(* IEC 61131-3 sources: plc-st-coding-agent/progress/evidence/f14_v3_parallel_20261112/jobs/codex_minimax-m27 (part 3) *)

(* ---- self-hard-01.raw_candidate_02.st ---- *)
FUNCTION_BLOCK FB
VAR_INPUT
    flowLow   : BOOL;
    ackBtn    : BOOL;
    sensorOK  : BOOL;
END_VAR
VAR_OUTPUT
    alarmActive : BOOL;
    alarmAcked  : BOOL;
    highHigh    : BOOL;
END_VAR
VAR
    prev_flowLow : BOOL := FALSE;
    prev_ackBtn  : BOOL := FALSE;
END_VAR

VAR_TEMP
    risingAck : BOOL;
END_VAR

risingAck := ackBtn AND NOT prev_ackBtn;

IF flowLow THEN
    // Condition is active
    IF NOT alarmActive THEN
        // New alarm activation
        alarmActive := TRUE;
        alarmAcked  := FALSE;
    ELSIF risingAck THEN
        // Rising ack while condition still exists - just mark acknowledged
        alarmAcked := TRUE;
    END_IF;
ELSE
    // Condition has disappeared
    IF prev_flowLow AND alarmAcked THEN
        // Condition just cleared, was already acknowledged - clear immediately
        alarmActive := FALSE;
        alarmAcked  := FALSE;
    ELSIF prev_flowLow AND NOT alarmAcked THEN
        // Condition just cleared, unacknowledged - enter pending clear state
        alarmAcked := TRUE;
    ELSIF risingAck AND alarmAcked THEN
        // Condition still gone from before, pending clear - clear on new ack
        alarmActive := FALSE;
        alarmAcked  := FALSE;
    END_IF;
END_IF;

// High priority alarm: sensor failure (independent)
highHigh := NOT sensorOK;

// Update state for next cycle
prev_flowLow := flowLow;
prev_ackBtn  := ackBtn;

END_FUNCTION_BLOCK

(* ---- self-hard-02.candidate_01.st ---- *)
FUNCTION_BLOCK FB
VAR_INPUT
    startBtn    : BOOL;
    abortBtn    : BOOL;
    setpoint    : REAL;
    pv          : REAL;
    maxDuration : INT;
END_VAR
VAR_OUTPUT
    elapsed : INT := 0;
    phase   : INT := 0;
    timeout : BOOL := FALSE;
END_VAR
VAR
    prev_startBtn : BOOL := FALSE;
    prev_phase    : INT  := 0;
    prev_elapsed  : INT  := 0;
    prev_timeout  : BOOL := FALSE;
END_VAR

// Priority 1: Abort (highest)
IF abortBtn THEN
    phase   := 9;
    elapsed := prev_elapsed;
    timeout := prev_timeout;

// Priority 2: New start rising edge (no abort)
ELSIF startBtn AND NOT prev_startBtn THEN
    phase   := 1;
    elapsed := 0;
    timeout := FALSE;

// Priority 3: Running states (prev phase 1 or 2)
ELSIF prev_phase = 1 OR prev_phase = 2 THEN
    elapsed := prev_elapsed + 1;

    IF elapsed >= maxDuration THEN
        timeout := TRUE;
        phase   := 3;
    ELSIF prev_phase = 1 AND pv >= setpoint THEN
        phase := 2;
    ELSE
        phase := prev_phase;
    END_IF;

// Priority 4: Frozen states (phase 0, 3, 9)
ELSE
    phase   := prev_phase;
    elapsed := prev_elapsed;
    timeout := prev_timeout;
END_IF;

prev_startBtn := startBtn;
prev_phase    := phase;
prev_elapsed  := elapsed;
prev_timeout  := timeout;
END_FUNCTION_BLOCK

(* ---- self-hard-02.raw_candidate_01.st ---- *)
FUNCTION_BLOCK FB
VAR_INPUT
    startBtn    : BOOL;
    abortBtn    : BOOL;
    setpoint    : REAL;
    pv          : REAL;
    maxDuration : INT;
END_VAR
VAR_OUTPUT
    elapsed : INT := 0;
    phase   : INT := 0;
    timeout : BOOL := FALSE;
END_VAR
VAR
    prev_startBtn : BOOL := FALSE;
    prev_phase    : INT  := 0;
    prev_elapsed  : INT  := 0;
    prev_timeout  : BOOL := FALSE;
END_VAR

// Priority 1: Abort (highest)
IF abortBtn THEN
    phase   := 9;
    elapsed := prev_elapsed;
    timeout := prev_timeout;

// Priority 2: New start rising edge (no abort)
ELSIF startBtn AND NOT prev_startBtn THEN
    phase   := 1;
    elapsed := 0;
    timeout := FALSE;

// Priority 3: Running states (prev phase 1 or 2)
ELSIF prev_phase = 1 OR prev_phase = 2 THEN
    elapsed := prev_elapsed + 1;

    IF elapsed >= maxDuration THEN
        timeout := TRUE;
        phase   := 3;
    ELSIF prev_phase = 1 AND pv >= setpoint THEN
        phase := 2;
    ELSE
        phase := prev_phase;
    END_IF;

// Priority 4: Frozen states (phase 0, 3, 9)
ELSE
    phase   := prev_phase;
    elapsed := prev_elapsed;
    timeout := prev_timeout;
END_IF;

prev_startBtn := startBtn;
prev_phase    := phase;
prev_elapsed  := elapsed;
prev_timeout  := timeout;
END_FUNCTION_BLOCK

(* ---- self-hard-03.candidate_01.st ---- *)
FUNCTION_BLOCK FB
VAR_INPUT
    pushEn: BOOL;
    pushItem: INT;
    popEn: BOOL;
END_VAR

VAR_IN_OUT
    fifo: ARRAY[1..8] OF INT;
END_VAR

VAR_OUTPUT
    count: INT := 0;
    full: BOOL := FALSE;
    empty: BOOL := TRUE;
    head: INT := 0;
END_VAR

VAR
    prevPushEn: BOOL := FALSE;
    prevPopEn: BOOL := FALSE;
END_VAR

VAR
    risingPush: BOOL;
    risingPop: BOOL;
    i: INT;
END_VAR

// Detect rising edges
risingPush := pushEn AND NOT prevPushEn;
risingPop := popEn AND NOT prevPopEn;

// Process in order: pop first, then push
// POP: only if queue not empty
IF risingPop AND count > 0 THEN
    // Shift left if more than one element
    IF count > 1 THEN
        FOR i := 1 TO count - 1 DO
            fifo[i] := fifo[i + 1];
        END_FOR;
    END_IF;
    // Decrement count
    count := count - 1;
END_IF;

// PUSH: only if queue not full
IF risingPush AND count < 8 THEN
    count := count + 1;
    fifo[count] := pushItem;
END_IF;

// Update outputs
full := (count = 8);
empty := (count = 0);
IF count > 0 THEN
    head := fifo[1];
ELSE
    head := 0;
END_IF;

// Save current state for next cycle
prevPushEn := pushEn;
prevPopEn := popEn;

END_FUNCTION_BLOCK

(* ---- self-hard-03.raw_candidate_01.st ---- *)
FUNCTION_BLOCK FB
VAR_INPUT
    pushEn: BOOL;
    pushItem: INT;
    popEn: BOOL;
END_VAR

VAR_IN_OUT
    fifo: ARRAY[1..8] OF INT;
END_VAR

VAR_OUTPUT
    count: INT := 0;
    full: BOOL := FALSE;
    empty: BOOL := TRUE;
    head: INT := 0;
END_VAR

VAR
    prevPushEn: BOOL := FALSE;
    prevPopEn: BOOL := FALSE;
END_VAR

VAR
    risingPush: BOOL;
    risingPop: BOOL;
    i: INT;
END_VAR

// Detect rising edges
risingPush := pushEn AND NOT prevPushEn;
risingPop := popEn AND NOT prevPopEn;

// Process in order: pop first, then push
// POP: only if queue not empty
IF risingPop AND count > 0 THEN
    // Shift left if more than one element
    IF count > 1 THEN
        FOR i := 1 TO count - 1 DO
            fifo[i] := fifo[i + 1];
        END_FOR;
    END_IF;
    // Decrement count
    count := count - 1;
END_IF;

// PUSH: only if queue not full
IF risingPush AND count < 8 THEN
    count := count + 1;
    fifo[count] := pushItem;
END_IF;

// Update outputs
full := (count = 8);
empty := (count = 0);
IF count > 0 THEN
    head := fifo[1];
ELSE
    head := 0;
END_IF;

// Save current state for next cycle
prevPushEn := pushEn;
prevPopEn := popEn;

END_FUNCTION_BLOCK

(* ---- self-hard-04.candidate_01.st ---- *)
FUNCTION_BLOCK FB
VAR
    prevDemand: INT := 0;
    prevLeadPump: INT := 0;
    prevRunningCount: INT := 0;
    prevLagPump: INT := 0;
    leadPump: INT := 0;
    lagPump: INT := 0;
    runningCount: INT := 0;
    minHours: LINT;
    minPumpIdx: INT;
    secondMinHours: LINT;
    secondMinIdx: INT;
    hoursDiff: LINT;
    needInitialLead: BOOL;
    needSwitchLead: BOOL;
    needRefreshLag: BOOL;
    i: INT;
    h: LINT;
END_VAR

// Clip demand to 0..5
IF demand < 0 THEN
    runningCount := 0;
ELSIF demand > 5 THEN
    runningCount := 5;
ELSE
    runningCount := demand;
END_IF;

// Detect state transitions
needInitialLead := (prevDemand = 0) AND (runningCount > 0);
needRefreshLag := (runningCount > prevRunningCount) OR (leadPump <> prevLeadPump);

// Find pump with minimum (runHours, pumpIdx)
minHours := runHours[1];
minPumpIdx := 1;
FOR i := 2 TO 5 DO
    h := runHours[i];
    IF (h < minHours) OR ((h = minHours) AND (i < minPumpIdx)) THEN
        minHours := h;
        minPumpIdx := i;
    END_IF;
END_FOR;

// Lead pump hysteresis check
IF leadPump >= 1 AND leadPump <= 5 THEN
    hoursDiff := runHours[leadPump] - minHours;
ELSE
    hoursDiff := 0;
END_IF;
needSwitchLead := (prevLeadPump <> 0) AND rotated AND (hoursDiff > 50);

// Demand = 0: clear both pumps immediately
IF runningCount = 0 THEN
    leadPump := 0;
    lagPump := 0;
    needRefreshLag := FALSE;
    needSwitchLead := FALSE;
END_IF;

// Handle lead pump change
IF needSwitchLead THEN
    leadPump := minPumpIdx;
    needRefreshLag := TRUE;
ELSIF needInitialLead THEN
    leadPump := minPumpIdx;
END_IF;

// Lag pump selection
IF needRefreshLag AND runningCount > 0 THEN
    secondMinHours := 16#7FFFFFFFFFFFFFFF;
    secondMinIdx := 0;
    FOR i := 1 TO 5 DO
        IF i <> leadPump THEN
            h := runHours[i];
            IF (h < secondMinHours) OR ((h = secondMinHours) AND (i < secondMinIdx)) THEN
                secondMinHours := h;
                secondMinIdx := i;
            END_IF;
        END_IF;
    END_FOR;
    lagPump := secondMinIdx;
ELSIF runningCount = 1 THEN
    lagPump := 0;
END_IF;

// Preserve lead pump if no change occurred
IF NOT needSwitchLead AND NOT needInitialLead AND runningCount > 0 THEN
    leadPump := prevLeadPump;
END_IF;

// Update previous-cycle state
prevDemand := runningCount;
prevLeadPump := leadPump;
prevRunningCount := runningCount;
prevLagPump := lagPump;

END_FUNCTION_BLOCK

(* ---- self-hard-04.candidate_02.st ---- *)
FUNCTION_BLOCK FB
VAR_INPUT
    demand: INT;
    runHours: ARRAY[1..5] OF LINT;
    rotated: BOOL;
END_VAR
VAR_OUTPUT
    leadPump: INT;
    lagPump: INT;
    runningCount: INT;
END_VAR
VAR
    prevDemand: INT := 0;
    prevLeadPump: INT := 0;
    prevRunningCount: INT := 0;
    prevLagPump: INT := 0;
    minHours: LINT;
    minPumpIdx: INT;
    secondMinHours: LINT;
    secondMinIdx: INT;
    hoursDiff: LINT;
    needInitialLead: BOOL;
    needSwitchLead: BOOL;
    needRefreshLag: BOOL;
    i: INT;
    h: LINT;
    clippedDemand: INT;
END_VAR

clippedDemand := demand;
IF clippedDemand < 0 THEN
    clippedDemand := 0;
ELSIF clippedDemand > 5 THEN
    clippedDemand := 5;
END_IF;

runningCount := clippedDemand;

needInitialLead := (prevDemand = 0) AND (runningCount > 0);
needRefreshLag := (runningCount > prevRunningCount) OR (leadPump <> prevLeadPump);

minHours := runHours[1];
minPumpIdx := 1;
FOR i := 2 TO 5 DO
    h := runHours[i];
    IF (h < minHours) OR ((h = minHours) AND (i < minPumpIdx)) THEN
        minHours := h;
        minPumpIdx := i;
    END_IF;
END_FOR;

IF leadPump >= 1 AND leadPump <= 5 THEN
    hoursDiff := runHours[leadPump] - minHours;
ELSE
    hoursDiff := 0;
END_IF;

needSwitchLead := (prevLeadPump <> 0) AND rotated AND (hoursDiff > 50);

IF runningCount = 0 THEN
    leadPump := 0;
    lagPump := 0;
ELSIF needSwitchLead THEN
    leadPump := minPumpIdx;
ELSIF needInitialLead THEN
    leadPump := minPumpIdx;
ELSE
    leadPump := prevLeadPump;
END_IF;

IF runningCount >= 2 THEN
    IF needRefreshLag THEN
        secondMinHours := 16#7FFFFFFFFFFFFFFF;
        secondMinIdx := 0;
        FOR i := 1 TO 5 DO
            IF i <> leadPump THEN
                h := runHours[i];
                IF (h < secondMinHours) OR ((h = secondMinHours) AND (i < secondMinIdx)) THEN
                    secondMinHours := h;
                    secondMinIdx := i;
                END_IF;
            END_IF;
        END_FOR;
        lagPump := secondMinIdx;
    ELSE
        lagPump := prevLagPump;
    END_IF;
ELSE
    lagPump := 0;
END_IF;

prevDemand := clippedDemand;
prevLeadPump := leadPump;
prevRunningCount := runningCount;
prevLagPump := lagPump;

END_FUNCTION_BLOCK

(* ---- self-hard-04.raw_candidate_01.st ---- *)
FUNCTION_BLOCK FB
VAR
    prevDemand: INT := 0;
    prevLeadPump: INT := 0;
    prevRunningCount: INT := 0;
    prevLagPump: INT := 0;
    leadPump: INT := 0;
    lagPump: INT := 0;
    runningCount: INT := 0;
    minHours: LINT;
    minPumpIdx: INT;
    secondMinHours: LINT;
    secondMinIdx: INT;
    hoursDiff: LINT;
    needInitialLead: BOOL;
    needSwitchLead: BOOL;
    needRefreshLag: BOOL;
    i: INT;
    h: LINT;
END_VAR

// Clip demand to 0..5
IF demand < 0 THEN
    runningCount := 0;
ELSIF demand > 5 THEN
    runningCount := 5;
ELSE
    runningCount := demand;
END_IF;

// Detect state transitions
needInitialLead := (prevDemand = 0) AND (runningCount > 0);
needRefreshLag := (runningCount > prevRunningCount) OR (leadPump <> prevLeadPump);

// Find pump with minimum (runHours, pumpIdx)
minHours := runHours[1];
minPumpIdx := 1;
FOR i := 2 TO 5 DO
    h := runHours[i];
    IF (h < minHours) OR ((h = minHours) AND (i < minPumpIdx)) THEN
        minHours := h;
        minPumpIdx := i;
    END_IF;
END_FOR;

// Lead pump hysteresis check
IF leadPump >= 1 AND leadPump <= 5 THEN
    hoursDiff := runHours[leadPump] - minHours;
ELSE
    hoursDiff := 0;
END_IF;
needSwitchLead := (prevLeadPump <> 0) AND rotated AND (hoursDiff > 50);

// Demand = 0: clear both pumps immediately
IF runningCount = 0 THEN
    leadPump := 0;
    lagPump := 0;
    needRefreshLag := FALSE;
    needSwitchLead := FALSE;
END_IF;

// Handle lead pump change
IF needSwitchLead THEN
    leadPump := minPumpIdx;
    needRefreshLag := TRUE;
ELSIF needInitialLead THEN
    leadPump := minPumpIdx;
END_IF;

// Lag pump selection
IF needRefreshLag AND runningCount > 0 THEN
    secondMinHours := 16#7FFFFFFFFFFFFFFF;
    secondMinIdx := 0;
    FOR i := 1 TO 5 DO
        IF i <> leadPump THEN
            h := runHours[i];
            IF (h < secondMinHours) OR ((h = secondMinHours) AND (i < secondMinIdx)) THEN
                secondMinHours := h;
                secondMinIdx := i;
            END_IF;
        END_IF;
    END_FOR;
    lagPump := secondMinIdx;
ELSIF runningCount = 1 THEN
    lagPump := 0;
END_IF;

// Preserve lead pump if no change occurred
IF NOT needSwitchLead AND NOT needInitialLead AND runningCount > 0 THEN
    leadPump := prevLeadPump;
END_IF;

// Update previous-cycle state
prevDemand := runningCount;
prevLeadPump := leadPump;
prevRunningCount := runningCount;
prevLagPump := lagPump;

END_FUNCTION_BLOCK

(* ---- self-hard-04.raw_candidate_02.st ---- *)
FUNCTION_BLOCK FB
VAR_INPUT
    demand: INT;
    runHours: ARRAY[1..5] OF LINT;
    rotated: BOOL;
END_VAR
VAR_OUTPUT
    leadPump: INT;
    lagPump: INT;
    runningCount: INT;
END_VAR
VAR
    prevDemand: INT := 0;
    prevLeadPump: INT := 0;
    prevRunningCount: INT := 0;
    prevLagPump: INT := 0;
    minHours: LINT;
    minPumpIdx: INT;
    secondMinHours: LINT;
    secondMinIdx: INT;
    hoursDiff: LINT;
    needInitialLead: BOOL;
    needSwitchLead: BOOL;
    needRefreshLag: BOOL;
    i: INT;
    h: LINT;
    clippedDemand: INT;
END_VAR

clippedDemand := demand;
IF clippedDemand < 0 THEN
    clippedDemand := 0;
ELSIF clippedDemand > 5 THEN
    clippedDemand := 5;
END_IF;

runningCount := clippedDemand;

needInitialLead := (prevDemand = 0) AND (runningCount > 0);
needRefreshLag := (runningCount > prevRunningCount) OR (leadPump <> prevLeadPump);

minHours := runHours[1];
minPumpIdx := 1;
FOR i := 2 TO 5 DO
    h := runHours[i];
    IF (h < minHours) OR ((h = minHours) AND (i < minPumpIdx)) THEN
        minHours := h;
        minPumpIdx := i;
    END_IF;
END_FOR;

IF leadPump >= 1 AND leadPump <= 5 THEN
    hoursDiff := runHours[leadPump] - minHours;
ELSE
    hoursDiff := 0;
END_IF;

needSwitchLead := (prevLeadPump <> 0) AND rotated AND (hoursDiff > 50);

IF runningCount = 0 THEN
    leadPump := 0;
    lagPump := 0;
ELSIF needSwitchLead THEN
    leadPump := minPumpIdx;
ELSIF needInitialLead THEN
    leadPump := minPumpIdx;
ELSE
    leadPump := prevLeadPump;
END_IF;

IF runningCount >= 2 THEN
    IF needRefreshLag THEN
        secondMinHours := 16#7FFFFFFFFFFFFFFF;
        secondMinIdx := 0;
        FOR i := 1 TO 5 DO
            IF i <> leadPump THEN
                h := runHours[i];
                IF (h < secondMinHours) OR ((h = secondMinHours) AND (i < secondMinIdx)) THEN
                    secondMinHours := h;
                    secondMinIdx := i;
                END_IF;
            END_IF;
        END_FOR;
        lagPump := secondMinIdx;
    ELSE
        lagPump := prevLagPump;
    END_IF;
ELSE
    lagPump := 0;
END_IF;

prevDemand := clippedDemand;
prevLeadPump := leadPump;
prevRunningCount := runningCount;
prevLagPump := lagPump;

END_FUNCTION_BLOCK

(* ---- self-hard-05.candidate_01.st ---- *)
FUNCTION_BLOCK FB
VAR_INPUT
    runRequest  : BOOL;
    flameOK     : BOOL;
    o2Valid     : BOOL;
    o2PV        : REAL;
    baseAir     : REAL;
    resetBtn    : BOOL;
END_VAR

VAR_OUTPUT
    fuelPermit  : BOOL;
    trimEnable  : BOOL;
    airTrim     : REAL;
    airCommand  : REAL;
    tripLatched : BOOL;
    o2Fault     : BOOL;
END_VAR

VAR
    prevResetBtn : BOOL := FALSE;
    tripInternal : BOOL := FALSE;
END_VAR

// 氧量故障判定
o2Fault := NOT o2Valid OR o2PV < 0.0 OR o2PV > 21.0;

// 熄火跳闸逻辑：运行中失去火焰当拍置位；安全停机态下复位上升沿清除
IF runRequest AND NOT flameOK THEN
    tripInternal := TRUE;
ELSIF NOT runRequest AND NOT flameOK AND resetBtn AND NOT prevResetBtn THEN
    tripInternal := FALSE;
END_IF;

// 燃料许可：运行请求、火焰正常、未跳闸三者同时成立
fuelPermit := runRequest AND flameOK AND NOT tripInternal;

// 氧量修正：投入需燃料许可且分析仪无故障
trimEnable := fuelPermit AND NOT o2Fault;
airTrim := 2.0 * (2.0 - o2PV);
airTrim := LIMIT(-10.0, airTrim, 10.0);
airTrim := SEL(trimEnable, 0.0, airTrim);

// 风门命令：基础开度叠加修正，偏置切除时自动归零
airCommand := baseAir + airTrim;
airCommand := LIMIT(0.0, airCommand, 100.0);
airCommand := SEL(fuelPermit, 0.0, airCommand);

// 输出跳闸状态
tripLatched := tripInternal;

// 边沿检测：保存复位按钮上一拍状态
prevResetBtn := resetBtn;

END_FUNCTION_BLOCK

(* ---- self-hard-05.candidate_02.st ---- *)
FUNCTION_BLOCK FB
VAR_INPUT
    runRequest  : BOOL;
    flameOK     : BOOL;
    o2Valid     : BOOL;
    o2PV        : REAL;
    baseAir     : REAL;
    resetBtn    : BOOL;
END_VAR

VAR_OUTPUT
    fuelPermit  : BOOL;
    trimEnable  : BOOL;
    airTrim     : REAL;
    airCommand  : REAL;
    tripLatched : BOOL;
    o2Fault     : BOOL;
END_VAR

VAR
    prevResetBtn : BOOL := FALSE;
    tripInternal : BOOL := FALSE;
END_VAR

// 氧量故障判定
o2Fault := NOT o2Valid OR o2PV < 0.0 OR o2PV > 21.0;

// 熄火跳闸逻辑：运行中失去火焰当拍置位；安全停机态下复位上升沿清除
IF runRequest AND NOT flameOK THEN
    tripInternal := TRUE;
ELSIF NOT runRequest AND NOT flameOK AND resetBtn AND NOT prevResetBtn THEN
    tripInternal := FALSE;
END_IF;

// 燃料许可：运行请求、火焰正常、未跳闸三者同时成立
fuelPermit := runRequest AND flameOK AND NOT tripInternal;

// 氧量修正：投入需燃料许可且分析仪无故障
IF fuelPermit AND NOT o2Fault THEN
    trimEnable := TRUE;
    airTrim := LIMIT(-10.0, 2.0 * (2.0 - o2PV), 10.0);
ELSE
    trimEnable := FALSE;
    airTrim := 0.0;
END_IF;

// 风门命令：基础开度叠加修正，偏置切除时自动归零
IF fuelPermit THEN
    airCommand := LIMIT(0.0, baseAir + airTrim, 100.0);
ELSE
    airCommand := 0.0;
END_IF;

// 输出跳闸状态
tripLatched := tripInternal;

// 边沿检测：保存复位按钮上一拍状态
prevResetBtn := resetBtn;

END_FUNCTION_BLOCK

(* ---- self-hard-05.raw_candidate_01.st ---- *)
FUNCTION_BLOCK FB
VAR_INPUT
    runRequest  : BOOL;
    flameOK     : BOOL;
    o2Valid     : BOOL;
    o2PV        : REAL;
    baseAir     : REAL;
    resetBtn    : BOOL;
END_VAR

VAR_OUTPUT
    fuelPermit  : BOOL;
    trimEnable  : BOOL;
    airTrim     : REAL;
    airCommand  : REAL;
    tripLatched : BOOL;
    o2Fault     : BOOL;
END_VAR

VAR
    prevResetBtn : BOOL := FALSE;
    tripInternal : BOOL := FALSE;
END_VAR

// 氧量故障判定
o2Fault := NOT o2Valid OR o2PV < 0.0 OR o2PV > 21.0;

// 熄火跳闸逻辑：运行中失去火焰当拍置位；安全停机态下复位上升沿清除
IF runRequest AND NOT flameOK THEN
    tripInternal := TRUE;
ELSIF NOT runRequest AND NOT flameOK AND resetBtn AND NOT prevResetBtn THEN
    tripInternal := FALSE;
END_IF;

// 燃料许可：运行请求、火焰正常、未跳闸三者同时成立
fuelPermit := runRequest AND flameOK AND NOT tripInternal;

// 氧量修正：投入需燃料许可且分析仪无故障
trimEnable := fuelPermit AND NOT o2Fault;
airTrim := 2.0 * (2.0 - o2PV);
airTrim := LIMIT(-10.0, airTrim, 10.0);
airTrim := SEL(trimEnable, 0.0, airTrim);

// 风门命令：基础开度叠加修正，偏置切除时自动归零
airCommand := baseAir + airTrim;
airCommand := LIMIT(0.0, airCommand, 100.0);
airCommand := SEL(fuelPermit, 0.0, airCommand);

// 输出跳闸状态
tripLatched := tripInternal;

// 边沿检测：保存复位按钮上一拍状态
prevResetBtn := resetBtn;

END_FUNCTION_BLOCK

(* ---- self-hard-05.raw_candidate_02.st ---- *)
FUNCTION_BLOCK FB
VAR_INPUT
    runRequest  : BOOL;
    flameOK     : BOOL;
    o2Valid     : BOOL;
    o2PV        : REAL;
    baseAir     : REAL;
    resetBtn    : BOOL;
END_VAR

VAR_OUTPUT
    fuelPermit  : BOOL;
    trimEnable  : BOOL;
    airTrim     : REAL;
    airCommand  : REAL;
    tripLatched : BOOL;
    o2Fault     : BOOL;
END_VAR

VAR
    prevResetBtn : BOOL := FALSE;
    tripInternal : BOOL := FALSE;
END_VAR

// 氧量故障判定
o2Fault := NOT o2Valid OR o2PV < 0.0 OR o2PV > 21.0;

// 熄火跳闸逻辑：运行中失去火焰当拍置位；安全停机态下复位上升沿清除
IF runRequest AND NOT flameOK THEN
    tripInternal := TRUE;
ELSIF NOT runRequest AND NOT flameOK AND resetBtn AND NOT prevResetBtn THEN
    tripInternal := FALSE;
END_IF;

// 燃料许可：运行请求、火焰正常、未跳闸三者同时成立
fuelPermit := runRequest AND flameOK AND NOT tripInternal;

// 氧量修正：投入需燃料许可且分析仪无故障
IF fuelPermit AND NOT o2Fault THEN
    trimEnable := TRUE;
    airTrim := LIMIT(-10.0, 2.0 * (2.0 - o2PV), 10.0);
ELSE
    trimEnable := FALSE;
    airTrim := 0.0;
END_IF;

// 风门命令：基础开度叠加修正，偏置切除时自动归零
IF fuelPermit THEN
    airCommand := LIMIT(0.0, baseAir + airTrim, 100.0);
ELSE
    airCommand := 0.0;
END_IF;

// 输出跳闸状态
tripLatched := tripInternal;

// 边沿检测：保存复位按钮上一拍状态
prevResetBtn := resetBtn;

END_FUNCTION_BLOCK

(* ---- self-hard-06.candidate_01.st ---- *)
FUNCTION_BLOCK FB
VAR_INPUT
    runRequest      : BOOL;
    pressure        : REAL;
    pressureValid   : BOOL;
    fuelFlow        : REAL;
    steamFlow       : REAL;
    outletCmd       : INT;
    outletFeedback  : INT;
    resetBtn        : BOOL;
END_VAR
VAR_OUTPUT
    tripLatched     : BOOL;
    fuelPermit      : BOOL;
    currentCauseMask: WORD;
    latchedCauseMask: WORD;
    diagnosticActive: BOOL;
END_VAR
VAR
    prevResetBtn    : BOOL := FALSE;
    stickyCounter   : INT  := 0;
END_VAR

// Reset edge detection
IF resetBtn AND NOT prevResetBtn THEN
    // Rising edge of reset button
    IF NOT runRequest AND pressureValid AND pressure <= 4200.0 THEN
        tripLatched     := FALSE;
        latchedCauseMask := 0;
    ELSE
        tripLatched := TRUE;
    END_IF;
ELSE
    // No reset edge
    IF tripLatched THEN
        tripLatched := TRUE;
    ELSIF runRequest AND (NOT pressureValid OR pressure >= 4500.0) THEN
        tripLatched := TRUE;
    END_IF;
END_IF;

// Valve sticking counter: reset on any interruption, increment only in valid overpressure
IF NOT runRequest OR NOT pressureValid OR pressure < 4500.0 OR outletCmd < 50 OR outletFeedback > 10 THEN
    stickyCounter := 0;
ELSIF outletCmd >= 50 AND outletFeedback <= 10 THEN
    stickyCounter := stickyCounter + 1;
END_IF;

// Determine current cause mask
currentCauseMask := 0;
IF runRequest THEN
    IF NOT pressureValid THEN
        currentCauseMask := 1;  // bit0 = 1
    ELSIF stickyCounter >= 3 THEN
        currentCauseMask := 2;  // bit1 = 2
    END_IF;

    IF pressureValid AND pressure >= 4500.0 THEN
        IF fuelFlow >= 4.0 AND steamFlow <= 10.0 THEN
            currentCauseMask := currentCauseMask OR 4;  // bit2 = 4
        END_IF;

        IF currentCauseMask = 0 THEN
            currentCauseMask := 8;  // bit3 = 8
        END_IF;
    END_IF;
END_IF;

// Accumulate latched mask during trip
IF tripLatched THEN
    latchedCauseMask := latchedCauseMask OR currentCauseMask;
END_IF;

// Outputs
fuelPermit      := runRequest AND NOT tripLatched;
diagnosticActive := (currentCauseMask <> 0);

// Update previous states
prevResetBtn := resetBtn;
END_FUNCTION_BLOCK

(* ---- self-hard-06.candidate_02.st ---- *)
FUNCTION_BLOCK FB
VAR_INPUT
    runRequest       : BOOL;
    pressure         : REAL;
    pressureValid    : BOOL;
    fuelFlow         : REAL;
    steamFlow        : REAL;
    outletCmd        : INT;
    outletFeedback   : INT;
    resetBtn         : BOOL;
END_VAR
VAR_OUTPUT
    tripLatched      : BOOL;
    fuelPermit       : BOOL;
    currentCauseMask : WORD;
    latchedCauseMask : WORD;
    diagnosticActive : BOOL;
END_VAR
VAR
    prevResetBtn     : BOOL := FALSE;
    stickyCounter    : INT  := 0;
END_VAR

// Rising edge detection for reset
VAR_TEMP
    resetRising : BOOL;
END_VAR
resetRising := resetBtn AND NOT prevResetBtn;

// S17 logic: latch holds from first trip until valid reset edge
IF resetRising AND NOT runRequest AND pressureValid AND pressure <= 4200.0 THEN
    tripLatched := FALSE;
    latchedCauseMask := 0;
ELSIF resetRising THEN
    tripLatched := TRUE;
    IF tripLatched THEN
        latchedCauseMask := latchedCauseMask OR currentCauseMask;
    END_IF;
ELSIF prevResetBtn OR tripLatched THEN
    tripLatched := TRUE;
    IF prevResetBtn OR tripLatched THEN
        latchedCauseMask := latchedCauseMask OR currentCauseMask;
    END_IF;
ELSIF runRequest AND (NOT pressureValid OR pressure >= 4500.0) THEN
    tripLatched := TRUE;
    latchedCauseMask := currentCauseMask;
ELSE
    tripLatched := FALSE;
END_IF;

// Valve sticking counter
IF NOT runRequest OR NOT pressureValid OR pressure < 4500.0 OR outletCmd < 50 OR outletFeedback > 10 THEN
    stickyCounter := 0;
ELSIF outletCmd >= 50 AND outletFeedback <= 10 THEN
    stickyCounter := stickyCounter + 1;
END_IF;

// Current cause mask
currentCauseMask := 0;
IF runRequest THEN
    IF NOT pressureValid THEN
        currentCauseMask := 1;
    ELSIF stickyCounter >= 3 THEN
        currentCauseMask := 2;
    END_IF;

    IF pressureValid AND pressure >= 4500.0 THEN
        IF fuelFlow >= 4.0 AND steamFlow <= 10.0 THEN
            currentCauseMask := currentCauseMask OR 4;
        END_IF;

        IF currentCauseMask = 0 THEN
            currentCauseMask := 8;
        END_IF;
    END_IF;
END_IF;

// Outputs
fuelPermit       := runRequest AND NOT tripLatched;
diagnosticActive := (currentCauseMask <> 0);

prevResetBtn := resetBtn;
END_FUNCTION_BLOCK

(* ---- self-hard-06.raw_candidate_01.st ---- *)
FUNCTION_BLOCK FB
VAR_INPUT
    runRequest      : BOOL;
    pressure        : REAL;
    pressureValid   : BOOL;
    fuelFlow        : REAL;
    steamFlow       : REAL;
    outletCmd       : INT;
    outletFeedback  : INT;
    resetBtn        : BOOL;
END_VAR
VAR_OUTPUT
    tripLatched     : BOOL;
    fuelPermit      : BOOL;
    currentCauseMask: WORD;
    latchedCauseMask: WORD;
    diagnosticActive: BOOL;
END_VAR
VAR
    prevResetBtn    : BOOL := FALSE;
    stickyCounter   : INT  := 0;
END_VAR

// Reset edge detection
IF resetBtn AND NOT prevResetBtn THEN
    // Rising edge of reset button
    IF NOT runRequest AND pressureValid AND pressure <= 4200.0 THEN
        tripLatched     := FALSE;
        latchedCauseMask := 0;
    ELSE
        tripLatched := TRUE;
    END_IF;
ELSE
    // No reset edge
    IF tripLatched THEN
        tripLatched := TRUE;
    ELSIF runRequest AND (NOT pressureValid OR pressure >= 4500.0) THEN
        tripLatched := TRUE;
    END_IF;
END_IF;

// Valve sticking counter: reset on any interruption, increment only in valid overpressure
IF NOT runRequest OR NOT pressureValid OR pressure < 4500.0 OR outletCmd < 50 OR outletFeedback > 10 THEN
    stickyCounter := 0;
ELSIF outletCmd >= 50 AND outletFeedback <= 10 THEN
    stickyCounter := stickyCounter + 1;
END_IF;

// Determine current cause mask
currentCauseMask := 0;
IF runRequest THEN
    IF NOT pressureValid THEN
        currentCauseMask := 1;  // bit0 = 1
    ELSIF stickyCounter >= 3 THEN
        currentCauseMask := 2;  // bit1 = 2
    END_IF;

    IF pressureValid AND pressure >= 4500.0 THEN
        IF fuelFlow >= 4.0 AND steamFlow <= 10.0 THEN
            currentCauseMask := currentCauseMask OR 4;  // bit2 = 4
        END_IF;

        IF currentCauseMask = 0 THEN
            currentCauseMask := 8;  // bit3 = 8
        END_IF;
    END_IF;
END_IF;

// Accumulate latched mask during trip
IF tripLatched THEN
    latchedCauseMask := latchedCauseMask OR currentCauseMask;
END_IF;

// Outputs
fuelPermit      := runRequest AND NOT tripLatched;
diagnosticActive := (currentCauseMask <> 0);

// Update previous states
prevResetBtn := resetBtn;
END_FUNCTION_BLOCK

(* ---- self-hard-06.raw_candidate_02.st ---- *)
FUNCTION_BLOCK FB
VAR_INPUT
    runRequest       : BOOL;
    pressure         : REAL;
    pressureValid    : BOOL;
    fuelFlow         : REAL;
    steamFlow        : REAL;
    outletCmd        : INT;
    outletFeedback   : INT;
    resetBtn         : BOOL;
END_VAR
VAR_OUTPUT
    tripLatched      : BOOL;
    fuelPermit       : BOOL;
    currentCauseMask : WORD;
    latchedCauseMask : WORD;
    diagnosticActive : BOOL;
END_VAR
VAR
    prevResetBtn     : BOOL := FALSE;
    stickyCounter    : INT  := 0;
END_VAR

// Rising edge detection for reset
VAR_TEMP
    resetRising : BOOL;
END_VAR
resetRising := resetBtn AND NOT prevResetBtn;

// S17 logic: latch holds from first trip until valid reset edge
IF resetRising AND NOT runRequest AND pressureValid AND pressure <= 4200.0 THEN
    tripLatched := FALSE;
    latchedCauseMask := 0;
ELSIF resetRising THEN
    tripLatched := TRUE;
    IF tripLatched THEN
        latchedCauseMask := latchedCauseMask OR currentCauseMask;
    END_IF;
ELSIF prevResetBtn OR tripLatched THEN
    tripLatched := TRUE;
    IF prevResetBtn OR tripLatched THEN
        latchedCauseMask := latchedCauseMask OR currentCauseMask;
    END_IF;
ELSIF runRequest AND (NOT pressureValid OR pressure >= 4500.0) THEN
    tripLatched := TRUE;
    latchedCauseMask := currentCauseMask;
ELSE
    tripLatched := FALSE;
END_IF;

// Valve sticking counter
IF NOT runRequest OR NOT pressureValid OR pressure < 4500.0 OR outletCmd < 50 OR outletFeedback > 10 THEN
    stickyCounter := 0;
ELSIF outletCmd >= 50 AND outletFeedback <= 10 THEN
    stickyCounter := stickyCounter + 1;
END_IF;

// Current cause mask
currentCauseMask := 0;
IF runRequest THEN
    IF NOT pressureValid THEN
        currentCauseMask := 1;
    ELSIF stickyCounter >= 3 THEN
        currentCauseMask := 2;
    END_IF;

    IF pressureValid AND pressure >= 4500.0 THEN
        IF fuelFlow >= 4.0 AND steamFlow <= 10.0 THEN
            currentCauseMask := currentCauseMask OR 4;
        END_IF;

        IF currentCauseMask = 0 THEN
            currentCauseMask := 8;
        END_IF;
    END_IF;
END_IF;

// Outputs
fuelPermit       := runRequest AND NOT tripLatched;
diagnosticActive := (currentCauseMask <> 0);

prevResetBtn := resetBtn;
END_FUNCTION_BLOCK

(* ---- self-hard-07.candidate_01.st ---- *)
FUNCTION_BLOCK FB
VAR_INPUT
    mode            : INT;
    resetBtn        : BOOL;
    scanSeconds     : REAL;
    tempSP          : REAL;
    tempPV          : REAL;
    flowPV          : REAL;
    manualFlowSP    : REAL;
    manualValve     : REAL;
END_VAR

VAR_OUTPUT
    flowSP          : REAL;
    valveCommand    : REAL;
    fault           : BOOL;
    normalMode      : BOOL;
END_VAR

VAR
    prevMode        : INT;
    prevResetBtn    : BOOL;
    prevFlowSP      : REAL;
    prevValveCmd    : REAL;
    prevTempSP      : REAL;
    accT            : REAL;
    accF            : REAL;
    firstScan       : BOOL;
END_VAR

fault := (mode < 0) OR (mode > 2) OR (scanSeconds <= 0.0) OR (scanSeconds > 10.0);

IF resetBtn AND NOT prevResetBtn THEN
    flowSP := manualFlowSP;
    valveCommand := manualValve;
    accT := 0.0;
    accF := 0.0;
    normalMode := FALSE;
    firstScan := FALSE;
    prevMode := mode;
    prevResetBtn := resetBtn;
    prevFlowSP := flowSP;
    prevValveCmd := valveCommand;
    prevTempSP := tempSP;
    RETURN;
END_IF;

IF mode <> prevMode THEN
    IF mode = 2 THEN
        flowSP := prevFlowSP;
        valveCommand := prevValveCmd;
    ELSE
        flowSP := manualFlowSP;
        valveCommand := prevValveCmd;
    END_IF;
    normalMode := FALSE;
    prevMode := mode;
    prevResetBtn := resetBtn;
    prevFlowSP := flowSP;
    prevValveCmd := valveCommand;
    prevTempSP := tempSP;
    RETURN;
END_IF;

IF firstScan THEN
    flowSP := manualFlowSP;
    valveCommand := manualValve;
    accT := 0.0;
    accF := 0.0;
    normalMode := FALSE;
    firstScan := FALSE;
    prevMode := mode;
    prevResetBtn := resetBtn;
    prevFlowSP := flowSP;
    prevValveCmd := valveCommand;
    prevTempSP := tempSP;
    RETURN;
END_IF;

normalMode := TRUE;

IF mode = 2 THEN
    VAR eF AT%Q* : REAL; END_VAR
    eF := flowSP - flowPV;
    accF := accF + 0.5 * eF * scanSeconds;
    valveCommand := 2.0 * eF + accF;
    valveCommand := LIMIT(0.0, valveCommand, 100.0);
    accF := valveCommand - 2.0 * eF;

    VAR eT AT%Q* : REAL; END_VAR
    eT := tempSP - tempPV;
    accT := accT + 0.2 * eT * scanSeconds;
    flowSP := 1.0 * eT + accT;
    flowSP := LIMIT(0.0, flowSP, 50.0);
    accT := flowSP - 1.0 * eT;
ELSIF mode = 1 THEN
    VAR eF AT%Q* : REAL; END_VAR
    eF := flowSP - flowPV;
    accF := accF + 0.5 * eF * scanSeconds;
    valveCommand := 2.0 * eF + accF;
    valveCommand := LIMIT(0.0, valveCommand, 100.0);
    accF := valveCommand - 2.0 * eF;
ELSE
    flowSP := manualFlowSP;
    valveCommand := manualValve;
END_IF;

prevMode := mode;
prevResetBtn := resetBtn;
prevFlowSP := flowSP;
prevValveCmd := valveCommand;
prevTempSP := tempSP;

END_FUNCTION_BLOCK

(* ---- self-hard-07.candidate_02.st ---- *)
FUNCTION_BLOCK FB
VAR_INPUT
    mode            : INT;
    resetBtn        : BOOL;
    scanSeconds     : REAL;
    tempSP          : REAL;
    tempPV          : REAL;
    flowPV          : REAL;
    manualFlowSP    : REAL;
    manualValve     : REAL;
END_VAR

VAR_OUTPUT
    flowSP          : REAL;
    valveCommand    : REAL;
    fault           : BOOL;
    normalMode      : BOOL;
END_VAR

VAR
    prevMode        : INT;
    prevResetBtn    : BOOL;
    prevFlowSP      : REAL;
    prevValveCmd    : REAL;
    accT            : REAL;
    accF            : REAL;
    firstScan       : BOOL;
    modeChanged     : BOOL;
END_VAR

    modeChanged := (mode <> prevMode);
    fault := (mode < 0) OR (mode > 2) OR (scanSeconds <= 0.0) OR (scanSeconds > 10.0);

    IF firstScan THEN
        flowSP := manualFlowSP;
        valveCommand := manualValve;
        accT := 0.0;
        accF := 0.0;
        normalMode := FALSE;
        firstScan := FALSE;
        prevMode := mode;
        prevResetBtn := resetBtn;
        prevFlowSP := flowSP;
        prevValveCmd := valveCommand;
        RETURN;
    END_IF;

    IF resetBtn AND NOT prevResetBtn THEN
        flowSP := manualFlowSP;
        valveCommand := manualValve;
        accT := 0.0;
        accF := 0.0;
        normalMode := FALSE;
        prevMode := mode;
        prevResetBtn := resetBtn;
        prevFlowSP := flowSP;
        prevValveCmd := valveCommand;
        RETURN;
    END_IF;

    IF fault THEN
        flowSP := manualFlowSP;
        valveCommand := manualValve;
        accT := 0.0;
        accF := 0.0;
        normalMode := FALSE;
        prevMode := mode;
        prevResetBtn := resetBtn;
        prevFlowSP := flowSP;
        prevValveCmd := valveCommand;
        RETURN;
    END_IF;

    IF modeChanged THEN
        IF mode = 2 THEN
            flowSP := prevFlowSP;
            valveCommand := prevValveCmd;
        ELSIF mode = 0 THEN
            flowSP := manualFlowSP;
            valveCommand := manualValve;
        ELSE
            flowSP := manualFlowSP;
            valveCommand := prevValveCmd;
        END_IF;
        normalMode := FALSE;
        prevMode := mode;
        prevResetBtn := resetBtn;
        prevFlowSP := flowSP;
        prevValveCmd := valveCommand;
        RETURN;
    END_IF;

    normalMode := TRUE;

    IF mode = 2 THEN
        accT := accT + 0.2 * (tempSP - tempPV) * scanSeconds;
        flowSP := 1.0 * (tempSP - tempPV) + accT;
        flowSP := LIMIT(0.0, flowSP, 50.0);
        accT := flowSP - 1.0 * (tempSP - tempPV);
        accF := accF + 0.5 * (flowSP - flowPV) * scanSeconds;
        valveCommand := 2.0 * (flowSP - flowPV) + accF;
        valveCommand := LIMIT(0.0, valveCommand, 100.0);
        accF := valveCommand - 2.0 * (flowSP - flowPV);
    ELSIF mode = 1 THEN
        flowSP := manualFlowSP;
        accF := accF + 0.5 * (flowSP - flowPV) * scanSeconds;
        valveCommand := 2.0 * (flowSP - flowPV) + accF;
        valveCommand := LIMIT(0.0, valveCommand, 100.0);
        accF := valveCommand - 2.0 * (flowSP - flowPV);
    ELSE
        flowSP := manualFlowSP;
        valveCommand := manualValve;
    END_IF;

    prevMode := mode;
    prevResetBtn := resetBtn;
    prevFlowSP := flowSP;
    prevValveCmd := valveCommand;

END_FUNCTION_BLOCK

(* ---- self-hard-07.raw_candidate_01.st ---- *)
FUNCTION_BLOCK FB
VAR_INPUT
    mode            : INT;
    resetBtn        : BOOL;
    scanSeconds     : REAL;
    tempSP          : REAL;
    tempPV          : REAL;
    flowPV          : REAL;
    manualFlowSP    : REAL;
    manualValve     : REAL;
END_VAR

VAR_OUTPUT
    flowSP          : REAL;
    valveCommand    : REAL;
    fault           : BOOL;
    normalMode      : BOOL;
END_VAR

VAR
    prevMode        : INT;
    prevResetBtn    : BOOL;
    prevFlowSP      : REAL;
    prevValveCmd    : REAL;
    prevTempSP      : REAL;
    accT            : REAL;
    accF            : REAL;
    firstScan       : BOOL;
END_VAR

fault := (mode < 0) OR (mode > 2) OR (scanSeconds <= 0.0) OR (scanSeconds > 10.0);

IF resetBtn AND NOT prevResetBtn THEN
    flowSP := manualFlowSP;
    valveCommand := manualValve;
    accT := 0.0;
    accF := 0.0;
    normalMode := FALSE;
    firstScan := FALSE;
    prevMode := mode;
    prevResetBtn := resetBtn;
    prevFlowSP := flowSP;
    prevValveCmd := valveCommand;
    prevTempSP := tempSP;
    RETURN;
END_IF

IF mode <> prevMode THEN
    IF mode = 2 THEN
        flowSP := prevFlowSP;
        valveCommand := prevValveCmd;
    ELSE
        flowSP := manualFlowSP;
        valveCommand := prevValveCmd;
    END_IF
    normalMode := FALSE;
    prevMode := mode;
    prevResetBtn := resetBtn;
    prevFlowSP := flowSP;
    prevValveCmd := valveCommand;
    prevTempSP := tempSP;
    RETURN;
END_IF

IF firstScan THEN
    flowSP := manualFlowSP;
    valveCommand := manualValve;
    accT := 0.0;
    accF := 0.0;
    normalMode := FALSE;
    firstScan := FALSE;
    prevMode := mode;
    prevResetBtn := resetBtn;
    prevFlowSP := flowSP;
    prevValveCmd := valveCommand;
    prevTempSP := tempSP;
    RETURN;
END_IF

normalMode := TRUE;

IF mode = 2 THEN
    VAR eF AT%Q* : REAL; END_VAR
    eF := flowSP - flowPV;
    accF := accF + 0.5 * eF * scanSeconds;
    valveCommand := 2.0 * eF + accF;
    valveCommand := LIMIT(0.0, valveCommand, 100.0);
    accF := valveCommand - 2.0 * eF;

    VAR eT AT%Q* : REAL; END_VAR
    eT := tempSP - tempPV;
    accT := accT + 0.2 * eT * scanSeconds;
    flowSP := 1.0 * eT + accT;
    flowSP := LIMIT(0.0, flowSP, 50.0);
    accT := flowSP - 1.0 * eT;
ELSIF mode = 1 THEN
    VAR eF AT%Q* : REAL; END_VAR
    eF := flowSP - flowPV;
    accF := accF + 0.5 * eF * scanSeconds;
    valveCommand := 2.0 * eF + accF;
    valveCommand := LIMIT(0.0, valveCommand, 100.0);
    accF := valveCommand - 2.0 * eF;
ELSE
    flowSP := manualFlowSP;
    valveCommand := manualValve;
END_IF;

prevMode := mode;
prevResetBtn := resetBtn;
prevFlowSP := flowSP;
prevValveCmd := valveCommand;
prevTempSP := tempSP;

END_FUNCTION_BLOCK

(* ---- self-hard-07.raw_candidate_02.st ---- *)
FUNCTION_BLOCK FB
VAR_INPUT
    mode            : INT;
    resetBtn        : BOOL;
    scanSeconds     : REAL;
    tempSP          : REAL;
    tempPV          : REAL;
    flowPV          : REAL;
    manualFlowSP    : REAL;
    manualValve     : REAL;
END_VAR

VAR_OUTPUT
    flowSP          : REAL;
    valveCommand    : REAL;
    fault           : BOOL;
    normalMode      : BOOL;
END_VAR

VAR
    prevMode        : INT;
    prevResetBtn    : BOOL;
    prevFlowSP      : REAL;
    prevValveCmd    : REAL;
    accT            : REAL;
    accF            : REAL;
    firstScan       : BOOL;
    modeChanged     : BOOL;
END_VAR

    modeChanged := (mode <> prevMode);
    fault := (mode < 0) OR (mode > 2) OR (scanSeconds <= 0.0) OR (scanSeconds > 10.0);

    IF firstScan THEN
        flowSP := manualFlowSP;
        valveCommand := manualValve;
        accT := 0.0;
        accF := 0.0;
        normalMode := FALSE;
        firstScan := FALSE;
        prevMode := mode;
        prevResetBtn := resetBtn;
        prevFlowSP := flowSP;
        prevValveCmd := valveCommand;
        RETURN;
    END_IF;

    IF resetBtn AND NOT prevResetBtn THEN
        flowSP := manualFlowSP;
        valveCommand := manualValve;
        accT := 0.0;
        accF := 0.0;
        normalMode := FALSE;
        prevMode := mode;
        prevResetBtn := resetBtn;
        prevFlowSP := flowSP;
        prevValveCmd := valveCommand;
        RETURN;
    END_IF;

    IF fault THEN
        flowSP := manualFlowSP;
        valveCommand := manualValve;
        accT := 0.0;
        accF := 0.0;
        normalMode := FALSE;
        prevMode := mode;
        prevResetBtn := resetBtn;
        prevFlowSP := flowSP;
        prevValveCmd := valveCommand;
        RETURN;
    END_IF;

    IF modeChanged THEN
        IF mode = 2 THEN
            flowSP := prevFlowSP;
            valveCommand := prevValveCmd;
        ELSIF mode = 0 THEN
            flowSP := manualFlowSP;
            valveCommand := manualValve;
        ELSE
            flowSP := manualFlowSP;
            valveCommand := prevValveCmd;
        END_IF;
        normalMode := FALSE;
        prevMode := mode;
        prevResetBtn := resetBtn;
        prevFlowSP := flowSP;
        prevValveCmd := valveCommand;
        RETURN;
    END_IF;

    normalMode := TRUE;

    IF mode = 2 THEN
        accT := accT + 0.2 * (tempSP - tempPV) * scanSeconds;
        flowSP := 1.0 * (tempSP - tempPV) + accT;
        flowSP := LIMIT(0.0, flowSP, 50.0);
        accT := flowSP - 1.0 * (tempSP - tempPV);
        accF := accF + 0.5 * (flowSP - flowPV) * scanSeconds;
        valveCommand := 2.0 * (flowSP - flowPV) + accF;
        valveCommand := LIMIT(0.0, valveCommand, 100.0);
        accF := valveCommand - 2.0 * (flowSP - flowPV);
    ELSIF mode = 1 THEN
        flowSP := manualFlowSP;
        accF := accF + 0.5 * (flowSP - flowPV) * scanSeconds;
        valveCommand := 2.0 * (flowSP - flowPV) + accF;
        valveCommand := LIMIT(0.0, valveCommand, 100.0);
        accF := valveCommand - 2.0 * (flowSP - flowPV);
    ELSE
        flowSP := manualFlowSP;
        valveCommand := manualValve;
    END_IF;

    prevMode := mode;
    prevResetBtn := resetBtn;
    prevFlowSP := flowSP;
    prevValveCmd := valveCommand;

END_FUNCTION_BLOCK

(* ---- self-medium-01.candidate_01.st ---- *)
FUNCTION_BLOCK FB
VAR_INPUT
    recipe      : ARRAY[1..8] OF ST_Recipe;
    selSlot     : INT;
    loadCmd     : BOOL;
    running     : BOOL;
END_VAR

VAR_OUTPUT
    valid       : BOOL;
    loadedID    : INT := 0;
END_VAR

VAR
    prevLoadCmd : BOOL := FALSE;
    prevValid   : BOOL := FALSE;
END_VAR

VAR_TEMP
    risingEdge  : BOOL;
BEGIN
    risingEdge := loadCmd AND NOT prevLoadCmd;

    IF running THEN
        // N10-S4: While running, hold state
        valid := prevValid;
        loadedID := 0;  // Will be overwritten by retention below
    ELSIF risingEdge THEN
        // Rising edge handling
        IF (selSlot >= 1) AND (selSlot <= 8) THEN
            // S5: Bounds check passed - safe to access array
            IF (recipe[selSlot].recipeID <> 0)
               AND (recipe[selSlot].totalRatio >= 99.0)
               AND (recipe[selSlot].totalRatio <= 101.0)
               AND (recipe[selSlot].temperature >= 30.0)
               AND (recipe[selSlot].temperature <= 180.0) THEN
                // All validations passed
                valid := TRUE;
                loadedID := recipe[selSlot].recipeID;
            ELSE
                // Validation failed
                valid := FALSE;
                loadedID := 0;
            END_IF;
        ELSE
            // S5: Slot out of bounds - invalid, no array access
            valid := FALSE;
            loadedID := 0;
        END_IF;
    ELSE
        // N10-S9: No rising edge - hold state
        valid := prevValid;
        loadedID := 0;  // Will be overwritten by retention below
    END_IF;

    // Retention when no rising edge or when running
    IF NOT risingEdge THEN
        loadedID := prevValid AND loadedID = 0 THEN 0 ELSE prevValid END_IF;
        IF running OR NOT risingEdge THEN
            loadedID := prevValid;  // Simplified retention
        END_IF;
    END_IF;

    prevValid := valid;
    prevLoadCmd := loadCmd;
END_FUNCTION_BLOCK

(* ---- self-medium-01.candidate_02.st ---- *)
TYPE ST_Recipe :
STRUCT
    recipeID    : INT;
    totalRatio  : REAL;
    temperature : REAL;
END_STRUCT;
END_TYPE;

FUNCTION_BLOCK FB
VAR_INPUT
    recipe      : ARRAY[1..8] OF ST_Recipe;
    selSlot     : INT;
    loadCmd     : BOOL;
    running     : BOOL;
END_VAR

VAR_OUTPUT
    valid       : BOOL := FALSE;
    loadedID    : INT := 0;
END_VAR

VAR
    prevLoadCmd : BOOL := FALSE;
    prevRunning : BOOL := FALSE;
END_VAR

BEGIN
    IF loadCmd AND NOT prevLoadCmd THEN
        IF NOT running THEN
            IF (selSlot >= 1) AND (selSlot <= 8) THEN
                IF (recipe[selSlot].recipeID <> 0) AND
                   (recipe[selSlot].totalRatio >= 99.0) AND
                   (recipe[selSlot].totalRatio <= 101.0) AND
                   (recipe[selSlot].temperature >= 30.0) AND
                   (recipe[selSlot].temperature <= 180.0) THEN
                    valid := TRUE;
                    loadedID := recipe[selSlot].recipeID;
                ELSE
                    valid := FALSE;
                    loadedID := 0;
                END_IF;
            ELSE
                valid := FALSE;
                loadedID := 0;
            END_IF;
        END_IF;
    END_IF;

    IF running AND NOT prevRunning THEN
        loadedID := loadedID;
    END_IF;

    prevLoadCmd := loadCmd;
    prevRunning := running;
END_FUNCTION_BLOCK

(* ---- self-medium-01.raw_candidate_01.st ---- *)
FUNCTION_BLOCK FB
VAR_INPUT
    recipe      : ARRAY[1..8] OF ST_Recipe;
    selSlot     : INT;
    loadCmd     : BOOL;
    running     : BOOL;
END_VAR

VAR_OUTPUT
    valid       : BOOL;
    loadedID    : INT := 0;
END_VAR

VAR
    prevLoadCmd : BOOL := FALSE;
    prevValid   : BOOL := FALSE;
END_VAR

VAR_TEMP
    risingEdge  : BOOL;
BEGIN
    risingEdge := loadCmd AND NOT prevLoadCmd;

    IF running THEN
        // N10-S4: While running, hold state
        valid := prevValid;
        loadedID := 0;  // Will be overwritten by retention below
    ELSIF risingEdge THEN
        // Rising edge handling
        IF (selSlot >= 1) AND (selSlot <= 8) THEN
            // S5: Bounds check passed - safe to access array
            IF (recipe[selSlot].recipeID <> 0)
               AND (recipe[selSlot].totalRatio >= 99.0)
               AND (recipe[selSlot].totalRatio <= 101.0)
               AND (recipe[selSlot].temperature >= 30.0)
               AND (recipe[selSlot].temperature <= 180.0) THEN
                // All validations passed
                valid := TRUE;
                loadedID := recipe[selSlot].recipeID;
            ELSE
                // Validation failed
                valid := FALSE;
                loadedID := 0;
            END_IF;
        ELSE
            // S5: Slot out of bounds - invalid, no array access
            valid := FALSE;
            loadedID := 0;
        END_IF;
    ELSE
        // N10-S9: No rising edge - hold state
        valid := prevValid;
        loadedID := 0;  // Will be overwritten by retention below
    END_IF;

    // Retention when no rising edge or when running
    IF NOT risingEdge THEN
        loadedID := prevValid AND loadedID = 0 THEN 0 ELSE prevValid END_IF;
        IF running OR NOT risingEdge THEN
            loadedID := prevValid;  // Simplified retention
        END_IF;
    END_IF;

    prevValid := valid;
    prevLoadCmd := loadCmd;
END_FUNCTION_BLOCK

(* ---- self-medium-01.raw_candidate_02.st ---- *)
TYPE ST_Recipe :
STRUCT
    recipeID    : INT;
    totalRatio  : REAL;
    temperature : REAL;
END_STRUCT
END_TYPE

FUNCTION_BLOCK FB
VAR_INPUT
    recipe      : ARRAY[1..8] OF ST_Recipe;
    selSlot     : INT;
    loadCmd     : BOOL;
    running     : BOOL;
END_VAR

VAR_OUTPUT
    valid       : BOOL := FALSE;
    loadedID    : INT := 0;
END_VAR

VAR
    prevLoadCmd : BOOL := FALSE;
    prevRunning : BOOL := FALSE;
END_VAR

BEGIN
    IF loadCmd AND NOT prevLoadCmd THEN
        IF NOT running THEN
            IF (selSlot >= 1) AND (selSlot <= 8) THEN
                IF (recipe[selSlot].recipeID <> 0) AND
                   (recipe[selSlot].totalRatio >= 99.0) AND
                   (recipe[selSlot].totalRatio <= 101.0) AND
                   (recipe[selSlot].temperature >= 30.0) AND
                   (recipe[selSlot].temperature <= 180.0) THEN
                    valid := TRUE;
                    loadedID := recipe[selSlot].recipeID;
                ELSE
                    valid := FALSE;
                    loadedID := 0;
                END_IF;
            ELSE
                valid := FALSE;
                loadedID := 0;
            END_IF;
        END_IF;
    END_IF;

    IF running AND NOT prevRunning THEN
        loadedID := loadedID;
    END_IF;

    prevLoadCmd := loadCmd;
    prevRunning := running;
END_FUNCTION_BLOCK

(* ---- self-medium-02.candidate_01.st ---- *)
FUNCTION_BLOCK FB
VAR
    buffer      : ARRAY[0..7] OF REAL;
    writeIndex  : INT := 0;
    sampleCount : INT := 0;
    windowFull  : BOOL := FALSE;
    sum         : REAL := 0.0;
END_VAR

VAR_INPUT
    enable   : BOOL;
    rawValue : REAL;
END_VAR

VAR_OUTPUT
    filteredValue : REAL := 0.0;
    windowFull    : BOOL := FALSE;
    sampleCount   : INT := 0;
END_VAR

BEGIN
    IF enable THEN
        // Determine index of oldest sample
        IF windowFull THEN
            // Buffer is full; oldest is at writeIndex
            sum := sum - buffer[writeIndex];
        ELSE
            // Buffer not full; oldest is at index 0
            IF sampleCount > 0 THEN
                sum := sum - buffer[0];
            END_IF;
        END_IF;

        // Add new sample
        sum := sum + rawValue;
        buffer[writeIndex] := rawValue;

        // Advance circular write pointer
        writeIndex := (writeIndex + 1) MOD 8;

        // Update sample count (cap at 8)
        IF sampleCount < 8 THEN
            sampleCount := sampleCount + 1;
        END_IF;

        // Update window full flag
        windowFull := (sampleCount = 8);

        // Compute arithmetic mean of valid samples
        IF sampleCount > 0 THEN
            filteredValue := sum / INT_TO_REAL(sampleCount);
        END_IF;
    ELSE
        // Enable is FALSE: clear all state
        sampleCount := 0;
        windowFull  := FALSE;
        writeIndex  := 0;
        sum         := 0.0;
        // filteredValue is NOT updated—holds last computed value
    END_IF;
END_FUNCTION_BLOCK

(* ---- self-medium-02.candidate_02.st ---- *)
FUNCTION_BLOCK FB
VAR_INPUT
    enable   : BOOL;
    rawValue : REAL;
END_VAR

VAR_OUTPUT
    filteredValue : REAL;
    windowFull    : BOOL;
    sampleCount   : INT;
END_VAR

VAR
    buffer     : ARRAY[0..7] OF REAL;
    writeIndex : INT := 0;
    sum        : REAL := 0.0;
END_VAR

BEGIN
    IF enable THEN
        IF windowFull THEN
            sum := sum - buffer[writeIndex];
        ELSIF sampleCount > 0 THEN
            sum := sum - buffer[0];
        END_IF;

        sum := sum + rawValue;
        buffer[writeIndex] := rawValue;
        writeIndex := (writeIndex + 1) MOD 8;

        IF sampleCount < 8 THEN
            sampleCount := sampleCount + 1;
        END_IF;

        windowFull := (sampleCount = 8);
        filteredValue := sum / INT_TO_REAL(sampleCount);
    ELSE
        sampleCount := 0;
        windowFull  := FALSE;
        writeIndex  := 0;
        sum         := 0.0;
    END_IF;
END_FUNCTION_BLOCK

(* ---- self-medium-02.raw_candidate_01.st ---- *)
FUNCTION_BLOCK FB
VAR
    buffer      : ARRAY[0..7] OF REAL;
    writeIndex  : INT := 0;
    sampleCount : INT := 0;
    windowFull  : BOOL := FALSE;
    sum         : REAL := 0.0;
END_VAR

VAR_INPUT
    enable   : BOOL;
    rawValue : REAL;
END_VAR

VAR_OUTPUT
    filteredValue : REAL := 0.0;
    windowFull    : BOOL := FALSE;
    sampleCount   : INT := 0;
END_VAR

BEGIN
    IF enable THEN
        // Determine index of oldest sample
        IF windowFull THEN
            // Buffer is full; oldest is at writeIndex
            sum := sum - buffer[writeIndex];
        ELSE
            // Buffer not full; oldest is at index 0
            IF sampleCount > 0 THEN
                sum := sum - buffer[0];
            END_IF;
        END_IF;

        // Add new sample
        sum := sum + rawValue;
        buffer[writeIndex] := rawValue;

        // Advance circular write pointer
        writeIndex := (writeIndex + 1) MOD 8;

        // Update sample count (cap at 8)
        IF sampleCount < 8 THEN
            sampleCount := sampleCount + 1;
        END_IF;

        // Update window full flag
        windowFull := (sampleCount = 8);

        // Compute arithmetic mean of valid samples
        IF sampleCount > 0 THEN
            filteredValue := sum / INT_TO_REAL(sampleCount);
        END_IF;
    ELSE
        // Enable is FALSE: clear all state
        sampleCount := 0;
        windowFull  := FALSE;
        writeIndex  := 0;
        sum         := 0.0;
        // filteredValue is NOT updated—holds last computed value
    END_IF;
END_FUNCTION_BLOCK

(* ---- self-medium-02.raw_candidate_02.st ---- *)
FUNCTION_BLOCK FB
VAR_INPUT
    enable   : BOOL;
    rawValue : REAL;
END_VAR

VAR_OUTPUT
    filteredValue : REAL;
    windowFull    : BOOL;
    sampleCount   : INT;
END_VAR

VAR
    buffer     : ARRAY[0..7] OF REAL;
    writeIndex : INT := 0;
    sum        : REAL := 0.0;
END_VAR

BEGIN
    IF enable THEN
        IF windowFull THEN
            sum := sum - buffer[writeIndex];
        ELSIF sampleCount > 0 THEN
            sum := sum - buffer[0];
        END_IF;

        sum := sum + rawValue;
        buffer[writeIndex] := rawValue;
        writeIndex := (writeIndex + 1) MOD 8;

        IF sampleCount < 8 THEN
            sampleCount := sampleCount + 1;
        END_IF;

        windowFull := (sampleCount = 8);
        filteredValue := sum / INT_TO_REAL(sampleCount);
    ELSE
        sampleCount := 0;
        windowFull  := FALSE;
        writeIndex  := 0;
        sum         := 0.0;
    END_IF;
END_FUNCTION_BLOCK

(* ---- self-medium-03.candidate_01.st ---- *)
FUNCTION_BLOCK FB
VAR_INPUT
    openBtn    : BOOL;
    closeBtn   : BOOL;
    openLimit  : BOOL;
    closeLimit : BOOL;
    obstacle   : BOOL;
END_VAR
VAR_OUTPUT
    motorUp    : BOOL := FALSE;
    motorDown  : BOOL := FALSE;
    errorFlag  : BOOL := FALSE;
END_VAR
VAR
    state       : UINT := 0;  // 0=IDLE, 1=OPENING, 2=CLOSING, 3=FAULT
    prevOpenBtn : BOOL := FALSE;
    prevCloseBtn: BOOL := FALSE;
END_VAR
VAR
    openBtnRising     : BOOL;
    closeBtnRising    : BOOL;
    bothBtnRising     : BOOL;
    prevBothBtn       : BOOL;
END_VAR

openBtnRising  := openBtn  AND NOT prevOpenBtn;
closeBtnRising := closeBtn AND NOT prevCloseBtn;
bothBtnRising  := (openBtn AND closeBtn) AND NOT prevBothBtn;

IF obstacle THEN
    state := FAULT;
    errorFlag := TRUE;
    motorUp   := FALSE;
    motorDown := FALSE;
ELSE
    CASE state OF
        0:  // IDLE
            motorUp   := FALSE;
            motorDown := FALSE;
            IF openBtnRising AND NOT closeBtn AND NOT openLimit THEN
                state := OPENING;
                motorUp := TRUE;
            ELSIF closeBtnRising AND NOT openBtn AND NOT closeLimit THEN
                state := CLOSING;
                motorDown := TRUE;
            END_IF;

        1:  // OPENING
            motorUp   := TRUE;
            motorDown := FALSE;
            IF openLimit THEN
                state := IDLE;
                motorUp := FALSE;
            END_IF;

        2:  // CLOSING
            motorUp   := FALSE;
            motorDown := TRUE;
            IF closeLimit THEN
                state := IDLE;
                motorDown := FALSE;
            END_IF;

        3:  // FAULT
            motorUp   := FALSE;
            motorDown := FALSE;
            IF bothBtnRising THEN
                state := IDLE;
            END_IF;
    END_CASE;
END_IF;

errorFlag      := (state = FAULT);
prevOpenBtn    := openBtn;
prevCloseBtn   := closeBtn;
prevBothBtn    := (openBtn AND closeBtn);

END_FUNCTION_BLOCK

(* ---- self-medium-03.candidate_02.st ---- *)
FUNCTION_BLOCK FB
VAR_INPUT
    openBtn    : BOOL;
    closeBtn   : BOOL;
    openLimit  : BOOL;
    closeLimit : BOOL;
    obstacle   : BOOL;
END_VAR
VAR_OUTPUT
    motorUp    : BOOL := FALSE;
    motorDown  : BOOL := FALSE;
    errorFlag  : BOOL := FALSE;
END_VAR
VAR
    state        : UINT := 0;
    prevOpenBtn  : BOOL := FALSE;
    prevCloseBtn : BOOL := FALSE;
    openBtnRising  : BOOL;
    closeBtnRising : BOOL;
    bothBtnRising  : BOOL;
END_VAR

openBtnRising  := openBtn  AND NOT prevOpenBtn;
closeBtnRising := closeBtn AND NOT prevCloseBtn;
bothBtnRising  := (openBtn AND closeBtn) AND (prevOpenBtn OR prevCloseBtn);

IF obstacle THEN
    state := 3;
    errorFlag := TRUE;
    motorUp   := FALSE;
    motorDown := FALSE;
ELSE
    CASE state OF
        0:  // IDLE
            motorUp   := FALSE;
            motorDown := FALSE;
            IF openBtnRising AND NOT closeBtn AND NOT openLimit THEN
                state := 1;
                motorUp := TRUE;
            ELSIF closeBtnRising AND NOT openBtn AND NOT closeLimit THEN
                state := 2;
                motorDown := TRUE;
            END_IF;

        1:  // OPENING
            motorUp   := TRUE;
            motorDown := FALSE;
            IF openLimit THEN
                state := 0;
                motorUp := FALSE;
            END_IF;

        2:  // CLOSING
            motorUp   := FALSE;
            motorDown := TRUE;
            IF closeLimit THEN
                state := 0;
                motorDown := FALSE;
            END_IF;

        3:  // FAULT
            motorUp   := FALSE;
            motorDown := FALSE;
            IF bothBtnRising THEN
                state := 0;
            END_IF;
    END_CASE;
END_IF;

errorFlag := (state = 3);
prevOpenBtn  := openBtn;
prevCloseBtn := closeBtn;

END_FUNCTION_BLOCK

(* ---- self-medium-03.raw_candidate_01.st ---- *)
FUNCTION_BLOCK FB
VAR_INPUT
    openBtn    : BOOL;
    closeBtn   : BOOL;
    openLimit  : BOOL;
    closeLimit : BOOL;
    obstacle   : BOOL;
END_VAR
VAR_OUTPUT
    motorUp    : BOOL := FALSE;
    motorDown  : BOOL := FALSE;
    errorFlag  : BOOL := FALSE;
END_VAR
VAR
    state       : UINT := 0;  // 0=IDLE, 1=OPENING, 2=CLOSING, 3=FAULT
    prevOpenBtn : BOOL := FALSE;
    prevCloseBtn: BOOL := FALSE;
END_VAR
VAR
    openBtnRising     : BOOL;
    closeBtnRising    : BOOL;
    bothBtnRising     : BOOL;
    prevBothBtn       : BOOL;
END_VAR

openBtnRising  := openBtn  AND NOT prevOpenBtn;
closeBtnRising := closeBtn AND NOT prevCloseBtn;
bothBtnRising  := (openBtn AND closeBtn) AND NOT prevBothBtn;

IF obstacle THEN
    state := FAULT;
    errorFlag := TRUE;
    motorUp   := FALSE;
    motorDown := FALSE;
ELSE
    CASE state OF
        0:  // IDLE
            motorUp   := FALSE;
            motorDown := FALSE;
            IF openBtnRising AND NOT closeBtn AND NOT openLimit THEN
                state := OPENING;
                motorUp := TRUE;
            ELSIF closeBtnRising AND NOT openBtn AND NOT closeLimit THEN
                state := CLOSING;
                motorDown := TRUE;
            END_IF

        1:  // OPENING
            motorUp   := TRUE;
            motorDown := FALSE;
            IF openLimit THEN
                state := IDLE;
                motorUp := FALSE;
            END_IF

        2:  // CLOSING
            motorUp   := FALSE;
            motorDown := TRUE;
            IF closeLimit THEN
                state := IDLE;
                motorDown := FALSE;
            END_IF

        3:  // FAULT
            motorUp   := FALSE;
            motorDown := FALSE;
            IF bothBtnRising THEN
                state := IDLE;
            END_IF
    END_CASE
END_IF;

errorFlag      := (state = FAULT);
prevOpenBtn    := openBtn;
prevCloseBtn   := closeBtn;
prevBothBtn    := (openBtn AND closeBtn);

END_FUNCTION_BLOCK

(* ---- self-medium-03.raw_candidate_02.st ---- *)
FUNCTION_BLOCK FB
VAR_INPUT
    openBtn    : BOOL;
    closeBtn   : BOOL;
    openLimit  : BOOL;
    closeLimit : BOOL;
    obstacle   : BOOL;
END_VAR
VAR_OUTPUT
    motorUp    : BOOL := FALSE;
    motorDown  : BOOL := FALSE;
    errorFlag  : BOOL := FALSE;
END_VAR
VAR
    state        : UINT := 0;
    prevOpenBtn  : BOOL := FALSE;
    prevCloseBtn : BOOL := FALSE;
    openBtnRising  : BOOL;
    closeBtnRising : BOOL;
    bothBtnRising  : BOOL;
END_VAR

openBtnRising  := openBtn  AND NOT prevOpenBtn;
closeBtnRising := closeBtn AND NOT prevCloseBtn;
bothBtnRising  := (openBtn AND closeBtn) AND (prevOpenBtn OR prevCloseBtn);

IF obstacle THEN
    state := 3;
    errorFlag := TRUE;
    motorUp   := FALSE;
    motorDown := FALSE;
ELSE
    CASE state OF
        0:  // IDLE
            motorUp   := FALSE;
            motorDown := FALSE;
            IF openBtnRising AND NOT closeBtn AND NOT openLimit THEN
                state := 1;
                motorUp := TRUE;
            ELSIF closeBtnRising AND NOT openBtn AND NOT closeLimit THEN
                state := 2;
                motorDown := TRUE;
            END_IF;

        1:  // OPENING
            motorUp   := TRUE;
            motorDown := FALSE;
            IF openLimit THEN
                state := 0;
                motorUp := FALSE;
            END_IF;

        2:  // CLOSING
            motorUp   := FALSE;
            motorDown := TRUE;
            IF closeLimit THEN
                state := 0;
                motorDown := FALSE;
            END_IF;

        3:  // FAULT
            motorUp   := FALSE;
            motorDown := FALSE;
            IF bothBtnRising THEN
                state := 0;
            END_IF;
    END_CASE;
END_IF;

errorFlag := (state = 3);
prevOpenBtn  := openBtn;
prevCloseBtn := closeBtn;

END_FUNCTION_BLOCK

(* ---- self-medium-04.candidate_01.st ---- *)
FUNCTION_BLOCK FB
VAR_INPUT
    startBtn    : BOOL;
    resetBtn    : BOOL;
    doneSensor  : BOOL;
    targetVol   : REAL;
    flowVol     : REAL;
END_VAR
VAR_OUTPUT
    valveOpen   : BOOL := FALSE;
    fillsToday  : INT := 0;
END_VAR
VAR
    prevStartBtn   : BOOL := FALSE;
    prevResetBtn   : BOOL := FALSE;
    prevValveOpen  : BOOL := FALSE;
    prevFillsToday : INT := 0;
    pending        : BOOL := FALSE;
    accumVol       : REAL := 0.0;
END_VAR

VAR
    risingStartBtn : BOOL;
    risingResetBtn : BOOL;
END_VAR

risingStartBtn := startBtn AND NOT prevStartBtn;
risingResetBtn := resetBtn AND NOT prevResetBtn;

prevFillsToday := fillsToday;
prevValveOpen  := valveOpen;

IF risingResetBtn THEN
    fillsToday := 0;
    pending    := FALSE;
    valveOpen  := FALSE;
    accumVol   := 0.0;
    prevFillsToday := 0;
    prevValveOpen  := FALSE;
ELSIF risingStartBtn THEN
    IF pending THEN
        pending := FALSE;
    END_IF;
    valveOpen := TRUE;
    accumVol  := 0.0;
ELSIF valveOpen THEN
    accumVol := accumVol + flowVol;
    IF accumVol >= targetVol THEN
        valveOpen := FALSE;
        pending   := TRUE;
    END_IF;
END_IF;

IF pending THEN
    IF doneSensor THEN
        IF prevFillsToday < 32767 THEN
            fillsToday := prevFillsToday + 1;
        ELSE
            fillsToday := 32767;
        END_IF;
        pending := FALSE;
    END_IF;
END_IF;

prevStartBtn  := startBtn;
prevResetBtn  := resetBtn;
END_FUNCTION_BLOCK

(* ---- self-medium-04.candidate_02.st ---- *)
FUNCTION_BLOCK FB
VAR_INPUT
    startBtn    : BOOL;
    resetBtn    : BOOL;
    doneSensor  : BOOL;
    targetVol   : REAL;
    flowVol     : REAL;
END_VAR
VAR_OUTPUT
    valveOpen   : BOOL := FALSE;
    fillsToday  : INT := 0;
END_VAR
VAR
    prevStartBtn   : BOOL := FALSE;
    prevResetBtn   : BOOL := FALSE;
    prevValveOpen  : BOOL := FALSE;
    prevFillsToday : INT := 0;
    pending        : BOOL := FALSE;
    accumVol       : REAL := 0.0;
END_VAR

VAR
    risingStartBtn : BOOL;
    risingResetBtn : BOOL;
END_VAR

risingStartBtn := startBtn AND NOT prevStartBtn;
risingResetBtn := resetBtn AND NOT prevResetBtn;
prevValveOpen  := valveOpen;
prevFillsToday := fillsToday;

IF risingResetBtn THEN
    fillsToday := 0;
    pending    := FALSE;
    valveOpen  := FALSE;
    accumVol   := 0.0;
    prevFillsToday := 0;
    prevValveOpen  := FALSE;
ELSIF risingStartBtn THEN
    IF pending THEN
        pending := FALSE;
    END_IF;
    IF prevValveOpen THEN
        accumVol := accumVol + flowVol;
    ELSE
        accumVol := flowVol;
    END_IF;
    IF accumVol >= targetVol THEN
        valveOpen := FALSE;
        pending   := TRUE;
    ELSE
        valveOpen := TRUE;
    END_IF;
ELSIF valveOpen THEN
    accumVol := accumVol + flowVol;
    IF accumVol >= targetVol THEN
        valveOpen := FALSE;
        pending   := TRUE;
    END_IF;
END_IF;

IF pending THEN
    IF doneSensor THEN
        IF prevFillsToday < 32767 THEN
            fillsToday := prevFillsToday + 1;
        ELSE
            fillsToday := 32767;
        END_IF;
        pending := FALSE;
    END_IF;
END_IF;

prevStartBtn  := startBtn;
prevResetBtn  := resetBtn;
END_FUNCTION_BLOCK

(* ---- self-medium-04.raw_candidate_01.st ---- *)
FUNCTION_BLOCK FB
VAR_INPUT
    startBtn    : BOOL;
    resetBtn    : BOOL;
    doneSensor  : BOOL;
    targetVol   : REAL;
    flowVol     : REAL;
END_VAR
VAR_OUTPUT
    valveOpen   : BOOL := FALSE;
    fillsToday  : INT := 0;
END_VAR
VAR
    prevStartBtn   : BOOL := FALSE;
    prevResetBtn   : BOOL := FALSE;
    prevValveOpen  : BOOL := FALSE;
    prevFillsToday : INT := 0;
    pending        : BOOL := FALSE;
    accumVol       : REAL := 0.0;
END_VAR

VAR
    risingStartBtn : BOOL;
    risingResetBtn : BOOL;
END_VAR

risingStartBtn := startBtn AND NOT prevStartBtn;
risingResetBtn := resetBtn AND NOT prevResetBtn;

prevFillsToday := fillsToday;
prevValveOpen  := valveOpen;

IF risingResetBtn THEN
    fillsToday := 0;
    pending    := FALSE;
    valveOpen  := FALSE;
    accumVol   := 0.0;
    prevFillsToday := 0;
    prevValveOpen  := FALSE;
ELSIF risingStartBtn THEN
    IF pending THEN
        pending := FALSE;
    END_IF;
    valveOpen := TRUE;
    accumVol  := 0.0;
ELSIF valveOpen THEN
    accumVol := accumVol + flowVol;
    IF accumVol >= targetVol THEN
        valveOpen := FALSE;
        pending   := TRUE;
    END_IF;
END_IF;

IF pending THEN
    IF doneSensor THEN
        IF prevFillsToday < 32767 THEN
            fillsToday := prevFillsToday + 1;
        ELSE
            fillsToday := 32767;
        END_IF;
        pending := FALSE;
    END_IF;
END_IF;

prevStartBtn  := startBtn;
prevResetBtn  := resetBtn;
END_FUNCTION_BLOCK

(* ---- self-medium-04.raw_candidate_02.st ---- *)
FUNCTION_BLOCK FB
VAR_INPUT
    startBtn    : BOOL;
    resetBtn    : BOOL;
    doneSensor  : BOOL;
    targetVol   : REAL;
    flowVol     : REAL;
END_VAR
VAR_OUTPUT
    valveOpen   : BOOL := FALSE;
    fillsToday  : INT := 0;
END_VAR
VAR
    prevStartBtn   : BOOL := FALSE;
    prevResetBtn   : BOOL := FALSE;
    prevValveOpen  : BOOL := FALSE;
    prevFillsToday : INT := 0;
    pending        : BOOL := FALSE;
    accumVol       : REAL := 0.0;
END_VAR

VAR
    risingStartBtn : BOOL;
    risingResetBtn : BOOL;
END_VAR

risingStartBtn := startBtn AND NOT prevStartBtn;
risingResetBtn := resetBtn AND NOT prevResetBtn;
prevValveOpen  := valveOpen;
prevFillsToday := fillsToday;

IF risingResetBtn THEN
    fillsToday := 0;
    pending    := FALSE;
    valveOpen  := FALSE;
    accumVol   := 0.0;
    prevFillsToday := 0;
    prevValveOpen  := FALSE;
ELSIF risingStartBtn THEN
    IF pending THEN
        pending := FALSE;
    END_IF;
    IF prevValveOpen THEN
        accumVol := accumVol + flowVol;
    ELSE
        accumVol := flowVol;
    END_IF;
    IF accumVol >= targetVol THEN
        valveOpen := FALSE;
        pending   := TRUE;
    ELSE
        valveOpen := TRUE;
    END_IF;
ELSIF valveOpen THEN
    accumVol := accumVol + flowVol;
    IF accumVol >= targetVol THEN
        valveOpen := FALSE;
        pending   := TRUE;
    END_IF;
END_IF;

IF pending THEN
    IF doneSensor THEN
        IF prevFillsToday < 32767 THEN
            fillsToday := prevFillsToday + 1;
        ELSE
            fillsToday := 32767;
        END_IF;
        pending := FALSE;
    END_IF;
END_IF;

prevStartBtn  := startBtn;
prevResetBtn  := resetBtn;
END_FUNCTION_BLOCK

(* ---- self-medium-05.candidate_01.st ---- *)
FUNCTION_BLOCK FB
VAR_INPUT
    enable       : BOOL;
    resetBtn     : BOOL;
    scanSeconds  : LREAL;
    steamFlow    : LREAL;
    fuelFlow     : LREAL;
    steamTemp    : LREAL;
    steamPressure: LREAL;
END_VAR

VAR_OUTPUT
    qualified   : BOOL;
    dataFault   : BOOL;
    qualifiedTon: LREAL;
    fuelTon     : LREAL;
    revenue     : LREAL;
    cost        : LREAL;
    netProfit   : LREAL;
END_VAR

VAR
    prevResetBtn : BOOL := FALSE;
END_VAR

VAR_TEMP
    resetRising : BOOL;
END_VAR

resetRising := resetBtn AND NOT prevResetBtn;

dataFault := (scanSeconds <= 0.0) OR (scanSeconds > 10.0)
    OR (steamFlow < 0.0) OR (steamFlow > 90.0)
    OR (fuelFlow < 0.0) OR (fuelFlow > 6.0);

qualified := (steamTemp >= 447.0) AND (steamTemp <= 453.0)
    AND (steamPressure >= 3750.0) AND (steamPressure <= 3850.0);

IF resetRising THEN
    qualifiedTon := 0.0;
    fuelTon := 0.0;
ELSIF enable AND NOT dataFault THEN
    fuelTon := fuelTon + fuelFlow * scanSeconds / 1000.0;
    IF qualified THEN
        qualifiedTon := qualifiedTon + steamFlow * scanSeconds / 1000.0;
    END_IF;
END_IF;

revenue := qualifiedTon * 280.0;
cost := fuelTon * 1500.0;
netProfit := revenue - cost;

prevResetBtn := resetBtn;

END_FUNCTION_BLOCK

(* ---- self-medium-05.raw_candidate_01.st ---- *)
FUNCTION_BLOCK FB
VAR_INPUT
    enable       : BOOL;
    resetBtn     : BOOL;
    scanSeconds  : LREAL;
    steamFlow    : LREAL;
    fuelFlow     : LREAL;
    steamTemp    : LREAL;
    steamPressure: LREAL;
END_VAR

VAR_OUTPUT
    qualified   : BOOL;
    dataFault   : BOOL;
    qualifiedTon: LREAL;
    fuelTon     : LREAL;
    revenue     : LREAL;
    cost        : LREAL;
    netProfit   : LREAL;
END_VAR

VAR
    prevResetBtn : BOOL := FALSE;
END_VAR

VAR_TEMP
    resetRising : BOOL;
END_VAR

resetRising := resetBtn AND NOT prevResetBtn;

dataFault := (scanSeconds <= 0.0) OR (scanSeconds > 10.0)
    OR (steamFlow < 0.0) OR (steamFlow > 90.0)
    OR (fuelFlow < 0.0) OR (fuelFlow > 6.0);

qualified := (steamTemp >= 447.0) AND (steamTemp <= 453.0)
    AND (steamPressure >= 3750.0) AND (steamPressure <= 3850.0);

IF resetRising THEN
    qualifiedTon := 0.0;
    fuelTon := 0.0;
ELSIF enable AND NOT dataFault THEN
    fuelTon := fuelTon + fuelFlow * scanSeconds / 1000.0;
    IF qualified THEN
        qualifiedTon := qualifiedTon + steamFlow * scanSeconds / 1000.0;
    END_IF;
END_IF;

revenue := qualifiedTon * 280.0;
cost := fuelTon * 1500.0;
netProfit := revenue - cost;

prevResetBtn := resetBtn;

END_FUNCTION_BLOCK

(* ---- self-medium-06.candidate_01.st ---- *)
FUNCTION_BLOCK FB
VAR_INPUT
    enable : BOOL;
    resetBtn : BOOL;
    sensorValid : BOOL;
    setpoint : REAL;
    temperature : REAL;
    scanSeconds : REAL;
    bias : REAL;
END_VAR

VAR_OUTPUT
    power : REAL := 0.0;
    correction : REAL := 0.0;
    fault : BOOL := FALSE;
END_VAR

VAR
    ePrev : REAL := 0.0;
    hasHistory : BOOL := FALSE;
    prevEnableAndNoFault : BOOL := FALSE;
    prevResetBtn : BOOL := FALSE;
END_VAR

VAR
    risingReset : BOOL;
    e : REAL;
    de : REAL;
    x : REAL;
    y : REAL;
    muNx : REAL;
    muZx : REAL;
    muPx : REAL;
    muNy : REAL;
    muZy : REAL;
    muPy : REAL;
    w1 : REAL;
    w2 : REAL;
    w3 : REAL;
    w4 : REAL;
    w5 : REAL;
    w6 : REAL;
    w7 : REAL;
    w8 : REAL;
    w9 : REAL;
    sumW : REAL;
    sumWc : REAL;
END_VAR

risingReset := resetBtn AND NOT prevResetBtn;
fault := NOT sensorValid OR scanSeconds <= 0.0 OR scanSeconds > 10.0;

IF fault OR risingReset OR NOT enable THEN
    ePrev := 0.0;
    hasHistory := FALSE;
END_IF;

IF scanSeconds <= 0.0 OR scanSeconds > 10.0 OR NOT sensorValid THEN
    power := 0.0;
    correction := 0.0;
    prevEnableAndNoFault := enable AND NOT fault;
    prevResetBtn := resetBtn;
    RETURN;
END_IF;

e := setpoint - temperature;

IF NOT hasHistory THEN
    de := 0.0;
ELSE
    de := (e - ePrev) / scanSeconds;
END_IF;

x := LIMIT(-1.0, e / 10.0, 1.0);
y := LIMIT(-1.0, de / 2.0, 1.0);

muNx := MAX(-x, 0.0);
muZx := 1.0 - ABS(x);
muPx := MAX(x, 0.0);

muNy := MAX(-y, 0.0);
muZy := 1.0 - ABS(y);
muPy := MAX(y, 0.0);

w1 := muNx * muNy;
w2 := muNx * muZy;
w3 := muNx * muPy;
w4 := muZx * muNy;
w5 := muZx * muZy;
w6 := muZx * muPy;
w7 := muPx * muNy;
w8 := muPx * muZy;
w9 := muPx * muPy;

sumW := w1 + w2 + w3 + w4 + w5 + w6 + w7 + w8 + w9;
sumWc := w1 * (-30.0) + w2 * (-20.0) + w3 * (-10.0) + w4 * (-10.0) + w5 * 0.0 + w6 * 10.0 + w7 * 10.0 + w8 * 20.0 + w9 * 30.0;

IF sumW > 0.0 THEN
    correction := sumWc / sumW;
ELSE
    correction := 0.0;
END_IF;

power := LIMIT(0.0, bias + correction, 100.0);

hasHistory := TRUE;
ePrev := e;
prevEnableAndNoFault := enable AND NOT fault;
prevResetBtn := resetBtn;
END_FUNCTION_BLOCK

(* ---- self-medium-06.candidate_02.st ---- *)
FUNCTION_BLOCK FB
VAR_INPUT
    enable : BOOL;
    resetBtn : BOOL;
    sensorValid : BOOL;
    setpoint : REAL;
    temperature : REAL;
    scanSeconds : REAL;
    bias : REAL;
END_VAR

VAR_OUTPUT
    power : REAL;
    correction : REAL;
    fault : BOOL;
END_VAR

VAR
    ePrev : REAL := 0.0;
    hasHistory : BOOL := FALSE;
    prevResetBtn : BOOL := FALSE;
END_VAR

VAR
    risingReset : BOOL;
    e : REAL;
    de : REAL;
    x : REAL;
    y : REAL;
    muNx : REAL;
    muZx : REAL;
    muPx : REAL;
    muNy : REAL;
    muZy : REAL;
    muPy : REAL;
    w1 : REAL;
    w2 : REAL;
    w3 : REAL;
    w4 : REAL;
    w5 : REAL;
    w6 : REAL;
    w7 : REAL;
    w8 : REAL;
    w9 : REAL;
    sumW : REAL;
    sumWc : REAL;
END_VAR

risingReset := resetBtn AND NOT prevResetBtn;
fault := NOT sensorValid OR scanSeconds <= 0.0 OR scanSeconds > 10.0;

IF fault OR risingReset THEN
    power := 0.0;
    correction := 0.0;
    ePrev := 0.0;
    hasHistory := FALSE;
END_IF;

IF NOT enable THEN
    power := 0.0;
    correction := 0.0;
END_IF;

IF NOT enable OR fault OR risingReset THEN
    prevResetBtn := resetBtn;
    RETURN;
END_IF;

e := setpoint - temperature;

IF NOT hasHistory THEN
    de := 0.0;
ELSE
    de := (e - ePrev) / scanSeconds;
END_IF;

x := LIMIT(-1.0, e / 10.0, 1.0);
y := LIMIT(-1.0, de / 2.0, 1.0);

muNx := MAX(-x, 0.0);
muZx := 1.0 - ABS(x);
muPx := MAX(x, 0.0);

muNy := MAX(-y, 0.0);
muZy := 1.0 - ABS(y);
muPy := MAX(y, 0.0);

w1 := muNx * muNy;
w2 := muNx * muZy;
w3 := muNx * muPy;
w4 := muZx * muNy;
w5 := muZx * muZy;
w6 := muZx * muPy;
w7 := muPx * muNy;
w8 := muPx * muZy;
w9 := muPx * muPy;

sumW := w1 + w2 + w3 + w4 + w5 + w6 + w7 + w8 + w9;
sumWc := w1 * (-30.0) + w2 * (-20.0) + w3 * (-10.0) + w4 * (-10.0) + w5 * 0.0 + w6 * 10.0 + w7 * 10.0 + w8 * 20.0 + w9 * 30.0;

IF sumW > 0.0 THEN
    correction := sumWc / sumW;
ELSE
    correction := 0.0;
END_IF;

power := LIMIT(0.0, bias + correction, 100.0);

hasHistory := TRUE;
ePrev := e;
prevResetBtn := resetBtn;
END_FUNCTION_BLOCK

(* ---- self-medium-06.raw_candidate_01.st ---- *)
FUNCTION_BLOCK FB
VAR_INPUT
    enable : BOOL;
    resetBtn : BOOL;
    sensorValid : BOOL;
    setpoint : REAL;
    temperature : REAL;
    scanSeconds : REAL;
    bias : REAL;
END_VAR

VAR_OUTPUT
    power : REAL := 0.0;
    correction : REAL := 0.0;
    fault : BOOL := FALSE;
END_VAR

VAR
    ePrev : REAL := 0.0;
    hasHistory : BOOL := FALSE;
    prevEnableAndNoFault : BOOL := FALSE;
    prevResetBtn : BOOL := FALSE;
END_VAR

VAR
    risingReset : BOOL;
    e : REAL;
    de : REAL;
    x : REAL;
    y : REAL;
    muNx : REAL;
    muZx : REAL;
    muPx : REAL;
    muNy : REAL;
    muZy : REAL;
    muPy : REAL;
    w1 : REAL;
    w2 : REAL;
    w3 : REAL;
    w4 : REAL;
    w5 : REAL;
    w6 : REAL;
    w7 : REAL;
    w8 : REAL;
    w9 : REAL;
    sumW : REAL;
    sumWc : REAL;
END_VAR

risingReset := resetBtn AND NOT prevResetBtn;
fault := NOT sensorValid OR scanSeconds <= 0.0 OR scanSeconds > 10.0;

IF fault OR risingReset OR NOT enable THEN
    ePrev := 0.0;
    hasHistory := FALSE;
END_IF;

IF scanSeconds <= 0.0 OR scanSeconds > 10.0 OR NOT sensorValid THEN
    power := 0.0;
    correction := 0.0;
    prevEnableAndNoFault := enable AND NOT fault;
    prevResetBtn := resetBtn;
    RETURN;
END_IF;

e := setpoint - temperature;

IF NOT hasHistory THEN
    de := 0.0;
ELSE
    de := (e - ePrev) / scanSeconds;
END_IF;

x := LIMIT(-1.0, e / 10.0, 1.0);
y := LIMIT(-1.0, de / 2.0, 1.0);

muNx := MAX(-x, 0.0);
muZx := 1.0 - ABS(x);
muPx := MAX(x, 0.0);

muNy := MAX(-y, 0.0);
muZy := 1.0 - ABS(y);
muPy := MAX(y, 0.0);

w1 := muNx * muNy;
w2 := muNx * muZy;
w3 := muNx * muPy;
w4 := muZx * muNy;
w5 := muZx * muZy;
w6 := muZx * muPy;
w7 := muPx * muNy;
w8 := muPx * muZy;
w9 := muPx * muPy;

sumW := w1 + w2 + w3 + w4 + w5 + w6 + w7 + w8 + w9;
sumWc := w1 * (-30.0) + w2 * (-20.0) + w3 * (-10.0) + w4 * (-10.0) + w5 * 0.0 + w6 * 10.0 + w7 * 10.0 + w8 * 20.0 + w9 * 30.0;

IF sumW > 0.0 THEN
    correction := sumWc / sumW;
ELSE
    correction := 0.0;
END_IF;

power := LIMIT(0.0, bias + correction, 100.0);

hasHistory := TRUE;
ePrev := e;
prevEnableAndNoFault := enable AND NOT fault;
prevResetBtn := resetBtn;
END_FUNCTION_BLOCK

(* ---- self-medium-06.raw_candidate_02.st ---- *)
FUNCTION_BLOCK FB
VAR_INPUT
    enable : BOOL;
    resetBtn : BOOL;
    sensorValid : BOOL;
    setpoint : REAL;
    temperature : REAL;
    scanSeconds : REAL;
    bias : REAL;
END_VAR

VAR_OUTPUT
    power : REAL;
    correction : REAL;
    fault : BOOL;
END_VAR

VAR
    ePrev : REAL := 0.0;
    hasHistory : BOOL := FALSE;
    prevResetBtn : BOOL := FALSE;
END_VAR

VAR
    risingReset : BOOL;
    e : REAL;
    de : REAL;
    x : REAL;
    y : REAL;
    muNx : REAL;
    muZx : REAL;
    muPx : REAL;
    muNy : REAL;
    muZy : REAL;
    muPy : REAL;
    w1 : REAL;
    w2 : REAL;
    w3 : REAL;
    w4 : REAL;
    w5 : REAL;
    w6 : REAL;
    w7 : REAL;
    w8 : REAL;
    w9 : REAL;
    sumW : REAL;
    sumWc : REAL;
END_VAR

risingReset := resetBtn AND NOT prevResetBtn;
fault := NOT sensorValid OR scanSeconds <= 0.0 OR scanSeconds > 10.0;

IF fault OR risingReset THEN
    power := 0.0;
    correction := 0.0;
    ePrev := 0.0;
    hasHistory := FALSE;
END_IF;

IF NOT enable THEN
    power := 0.0;
    correction := 0.0;
END_IF;

IF NOT enable OR fault OR risingReset THEN
    prevResetBtn := resetBtn;
    RETURN;
END_IF;

e := setpoint - temperature;

IF NOT hasHistory THEN
    de := 0.0;
ELSE
    de := (e - ePrev) / scanSeconds;
END_IF;

x := LIMIT(-1.0, e / 10.0, 1.0);
y := LIMIT(-1.0, de / 2.0, 1.0);

muNx := MAX(-x, 0.0);
muZx := 1.0 - ABS(x);
muPx := MAX(x, 0.0);

muNy := MAX(-y, 0.0);
muZy := 1.0 - ABS(y);
muPy := MAX(y, 0.0);

w1 := muNx * muNy;
w2 := muNx * muZy;
w3 := muNx * muPy;
w4 := muZx * muNy;
w5 := muZx * muZy;
w6 := muZx * muPy;
w7 := muPx * muNy;
w8 := muPx * muZy;
w9 := muPx * muPy;

sumW := w1 + w2 + w3 + w4 + w5 + w6 + w7 + w8 + w9;
sumWc := w1 * (-30.0) + w2 * (-20.0) + w3 * (-10.0) + w4 * (-10.0) + w5 * 0.0 + w6 * 10.0 + w7 * 10.0 + w8 * 20.0 + w9 * 30.0;

IF sumW > 0.0 THEN
    correction := sumWc / sumW;
ELSE
    correction := 0.0;
END_IF;

power := LIMIT(0.0, bias + correction, 100.0);

hasHistory := TRUE;
ePrev := e;
prevResetBtn := resetBtn;
END_FUNCTION_BLOCK
